// TIA Portal project "Project1" (V16)

(* hardware
DEVICE "S7300/ET200M station_1"  S7-300 station
   slot 0: "Rail_0"  Rail  6ES7 390-1***0-0AA0
   slot 2: "PLC_1"  CPU 315-2 DP  6ES7 315-2AG10-0AB0  V2.6
      slot 0: "MPI interface_1"  X1
      slot 1: "DP interface_1"  X2
*)

// ===== PLC "PLC_1"  CPU 315-2 DP =====

VAR_GLOBAL   // PLC tag table "Default tag table"
   "Tag_1" AT %MW10 : Word;
   "Tag_2" AT %MW20 : Word;
   "Tag_3" AT %M0.0 : Bool;
   "Tag_4" AT %M0.1 : Bool;
END_VAR

DATA_BLOCK "DB1"   // DB1
{ S7_Optimized_Access := 'FALSE' }
VERSION : 0.1
   VAR
      one : Int;
      one_1 : Int;
      one_2 : Int;
      one_3 : Int;
      one_4 : Int;
      one_5 : Int;
      one_6 : Int;
      one_7 : Int;
      one_1_1 : Int;
      one_2_1 : Int;
      one_3_1 : Int;
      one_4_1 : Int;
      one_5_1 : Int;
      one_5_2 : Int;
      one_5_3 : Int;
      one_5_4 : Int;
      one_5_5 : Int;
      one_5_6 : Int;
      one_5_7 : Int;
      one_5_8 : Int;
      one_5_9 : Int;
      one_5_10 : Int;
      one_5_11 : Int;
      one_5_12 : Int;
      one_5_13 : Int;
   END_VAR
BEGIN
END_DATA_BLOCK

DATA_BLOCK "DB2"   // DB2
{ S7_Optimized_Access := 'FALSE' }
VERSION : 0.1
   VAR
      Static_1 : Int;
      Static_2 : Int;
      Static_3 : Int;
      Static_4 : Int;
      Static_5 : Int;
      Static_6 : Int;
      Static_7 : Int;
      Static_8 : Int;
      Static_9 : Int;
      Static_10 : Int;
      Static_11 : Int;
      Static_12 : Int;
      Static_13 : Int;
      Static_14 : Int;
      Static_15 : Int;
      Static_16 : Int;
      Static_17 : Int;
      Static_18 : Int;
      Static_19 : Int;
      Static_20 : Int;
      Static_21 : Int;
      Static_22 : Int;
      Static_23 : Int;
      Static_24 : Int;
      Static_25 : Int;
   END_VAR
BEGIN
END_DATA_BLOCK

FUNCTION "FC1" : Void   // FC1, STL
{ S7_Optimized_Access := 'FALSE' }
VERSION : 0.1
BEGIN

REGION Network 1
         L     "Tag_1";
         L     "Tag_2";
         >I;
         S     "Tag_3";

         <I;
         S     "Tag_4";
END_REGION
END_FUNCTION

FUNCTION "FC2" : Void   // FC2, STL
{ S7_Optimized_Access := 'FALSE' }
VERSION : 0.1
BEGIN

REGION Network 1
         L     "DB1".one_5;
         L     "DB1".one_3_1;
         >I;
         S     "Tag_3";

         <I;
         S     "Tag_4";
END_REGION
END_FUNCTION

FUNCTION "FC3" : Void   // FC3, STL
{ S7_Optimized_Access := 'FALSE' }
VERSION : 0.1
BEGIN

REGION Network 1
         L     "DB2".Static_6;
         L     "DB2".Static_11;
         >I;
         S     "Tag_3";

         <I;
         S     "Tag_4";
END_REGION
END_FUNCTION

ORGANIZATION_BLOCK "Main"   // OB1, STL
TITLE = "Main Program Sweep (Cycle)"
{ S7_Optimized_Access := 'FALSE' }
VERSION : 0.1
   VAR_TEMP
      OB1_EV_CLASS : Byte;   // Bits 0-3 = 1 (Coming event), Bits 4-7 = 1 (Event class 1)
      OB1_SCAN_1 : Byte;   // 1 (Cold restart scan 1 of OB 1), 3 (Scan 2-n of OB 1)
      OB1_PRIORITY : Byte;   // Priority of OB Execution
      OB1_OB_NUMBR : Byte;   // 1 (Organization block 1, OB1)
      OB1_RESERVED_1 : Byte;   // Reserved for system
      OB1_RESERVED_2 : Byte;   // Reserved for system
      OB1_PREV_CYCLE : Int;   // Cycle time of previous OB1 scan (milliseconds)
      OB1_MIN_CYCLE : Int;   // Minimum cycle time of OB1 (milliseconds)
      OB1_MAX_CYCLE : Int;   // Maximum cycle time of OB1 (milliseconds)
      OB1_DATE_TIME : Date_And_Time;   // Date and time OB1 started
   END_VAR
BEGIN

REGION Network 1
   //CALL  "FC1"
   //  CALL  "FC2"
         CALL  "FC3";
END_REGION
END_ORGANIZATION_BLOCK